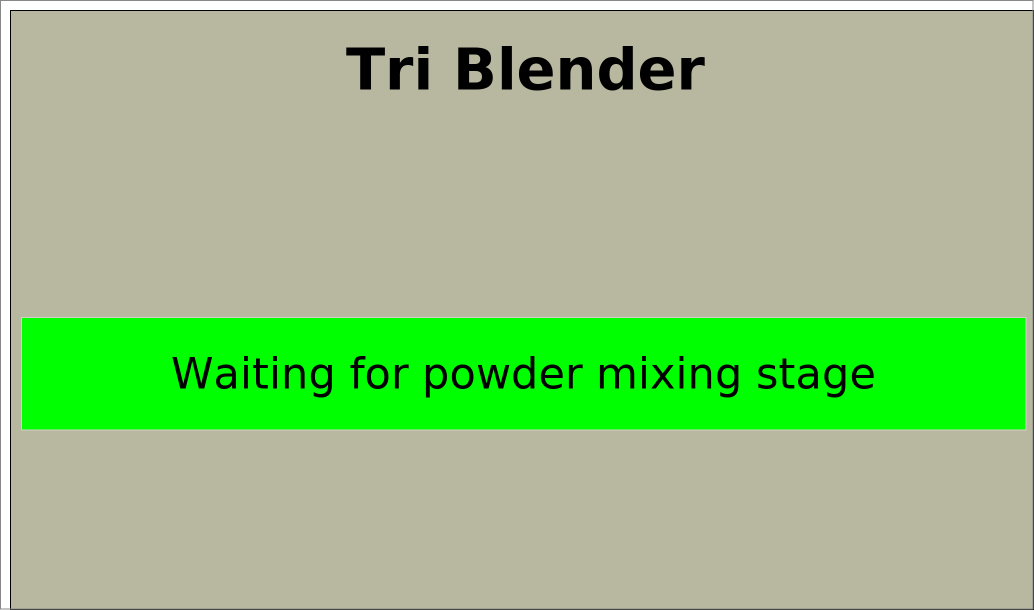
VISUALIZATION StartVisu  // 1034x610
    Rectangle (10,10 1024x600)
    Textfield (19,21 1013x96), "Tri Blender"
    Textfield (21,317 1005x113), "Waiting for powder mixing stage"
END_VISUALIZATION

(* stored: Version 1.1.0.1, ProductVersion 3.1.4024.12
   Visu StartVisu: Id {6004dca2-3ce1-443e-a6dd-2ca443b4e8e3} *)
